(* IEC 61131-3 sources: 2026_Projet_YGO_ExcavatriceDragage/TOOLS/TEST_AUTO_CI/RESULTS/B_AU_SECURITE/reports, 1 file *)

(* ---- FB_Safety_EmergencyManagement_test.st ---- *)
SETUP
VAR
    fb : FB_SAFETY_EMERGENCYMANAGEMENT;
END_VAR
END_SETUP

(* Profil actif : 12 preuves fonctionnelles AF. Les essais de causes et diagnostics sont conserves dans contract_deferred. *)

(* Ordre de rapport stable : contrat IEC, scenarios operationnels, puis TC-P01 par numero croissant. *)

TEST 'TC-P03-001 Dynamique Enable : neutralisation initiale, transition Ready au repos, puis coupure'
    (* Scan 0 : Enable=FALSE -> Neutralisation standard *)
    fb(ENABLE := FALSE, RESET := FALSE, ARMREQUEST := FALSE, POWERCUTOFFREQUEST := FALSE,
       BTNEMERGENCYCUTOFF := FALSE, EMERGENCYCHAINCLOSED := TRUE, POWERCONTACTORENGAGED := FALSE);
    fb(ENABLE := FALSE, RESET := FALSE, ARMREQUEST := FALSE, POWERCUTOFFREQUEST := FALSE,
       BTNEMERGENCYCUTOFF := FALSE, EMERGENCYCHAINCLOSED := TRUE, POWERCONTACTORENGAGED := FALSE);
    ASSERT_FALSE(fb.STATUS.READY, 'Enable=FALSE -> Ready=FALSE (neutralise)');
    ASSERT_FALSE(fb.STATUS.DIAG.ERROR, 'Enable=FALSE -> Pas d erreur');
    ASSERT_FALSE(fb.CMD.MAINTAINA_CMD, 'Enable=FALSE -> MaintainA_Cmd=FALSE (projection fail-safe §10)');
    ASSERT_FALSE(fb.CMD.MAINTAINB_CMD, 'Enable=FALSE -> MaintainB_Cmd=FALSE (projection fail-safe §10)');
    ASSERT_FALSE(fb.CMD.ARMPULSE_CMD, 'Enable=FALSE -> ArmPulse_Cmd=FALSE (projection fail-safe §10)');
    ASSERT_EQ(fb.STATUS.STATE.STEP, 0, 'Enable=FALSE -> sequence neutralisee, Step=0');
    ASSERT_EQ(fb.STATUS.OPERATORMESSAGE, 'AU neutralisee (Enable=FALSE)', 'message neutralisation (gate §2, priorite §11)');

    ADVANCE_TIME(10000000);

    (* Scan 1 : Enable=TRUE -> Prete en service *)
    fb(ENABLE := TRUE, RESET := FALSE, ARMREQUEST := FALSE, POWERCUTOFFREQUEST := FALSE,
       BTNEMERGENCYCUTOFF := FALSE, EMERGENCYCHAINCLOSED := TRUE, POWERCONTACTORENGAGED := FALSE);
    fb(ENABLE := TRUE, RESET := FALSE, ARMREQUEST := FALSE, POWERCUTOFFREQUEST := FALSE,
       BTNEMERGENCYCUTOFF := FALSE, EMERGENCYCHAINCLOSED := TRUE, POWERCONTACTORENGAGED := FALSE);
    ASSERT_TRUE(fb.STATUS.READY, 'Enable=TRUE -> Ready=TRUE (nominal)');
    ASSERT_FALSE(fb.STATUS.DIAG.ERROR, 'Au repos -> Pas d erreur');

    ADVANCE_TIME(10000000);

    (* Scan 2 : Enable=FALSE -> Re-neutralisation *)
    fb(ENABLE := FALSE, RESET := FALSE, ARMREQUEST := FALSE, POWERCUTOFFREQUEST := FALSE,
       BTNEMERGENCYCUTOFF := FALSE, EMERGENCYCHAINCLOSED := TRUE, POWERCONTACTORENGAGED := FALSE);
    fb(ENABLE := FALSE, RESET := FALSE, ARMREQUEST := FALSE, POWERCUTOFFREQUEST := FALSE,
       BTNEMERGENCYCUTOFF := FALSE, EMERGENCYCHAINCLOSED := TRUE, POWERCONTACTORENGAGED := FALSE);
    ASSERT_FALSE(fb.STATUS.READY, 'Coupure -> Ready retombe a FALSE');
END_TEST

TEST 'TC-P01-SCEN-NOM Scenario Nominal : Sequence complete de rearmement sans blocage'
    (* 💤 Étape 0 : Repos initial (machine hors tension, contacteur au repos, Armable=TRUE) *)
    fb(ENABLE := TRUE, RESET := FALSE, ARMREQUEST := FALSE, POWERCUTOFFREQUEST := FALSE,
       BTNEMERGENCYCUTOFF := FALSE, EMERGENCYCHAINCLOSED := TRUE, POWERCONTACTORENGAGED := FALSE);
    fb(ENABLE := TRUE, RESET := FALSE, ARMREQUEST := FALSE, POWERCUTOFFREQUEST := FALSE,
       BTNEMERGENCYCUTOFF := FALSE, EMERGENCYCHAINCLOSED := TRUE, POWERCONTACTORENGAGED := FALSE);
    ADVANCE_TIME(10000000);
    fb(ENABLE := TRUE, RESET := FALSE, ARMREQUEST := FALSE, POWERCUTOFFREQUEST := FALSE,
       BTNEMERGENCYCUTOFF := FALSE, EMERGENCYCHAINCLOSED := TRUE, POWERCONTACTORENGAGED := FALSE);
    fb(ENABLE := TRUE, RESET := FALSE, ARMREQUEST := FALSE, POWERCUTOFFREQUEST := FALSE,
       BTNEMERGENCYCUTOFF := FALSE, EMERGENCYCHAINCLOSED := TRUE, POWERCONTACTORENGAGED := FALSE);
    ASSERT_TRUE(fb.STATUS.STATE.ARMABLE, 'Au repos boucle saine -> Armable=TRUE');
    ASSERT_FALSE(fb.STATUS.DONE, 'Puissance non encore engagee -> Done=FALSE');
    ASSERT_EQ(fb.STATUS.OPERATORMESSAGE, 'AU: repos - pret a rearmer', 'message CASE 0/IDLE au repos sain');

    (* ⏱️ Étape 0bis : Demande de réarmement (Front ArmRequest -> Délai pré-armement 500ms en Step 0) *)
    ADVANCE_TIME(10000000);
    fb(ENABLE := TRUE, RESET := FALSE, ARMREQUEST := TRUE, POWERCUTOFFREQUEST := FALSE,
       BTNEMERGENCYCUTOFF := FALSE, EMERGENCYCHAINCLOSED := TRUE, POWERCONTACTORENGAGED := FALSE);
    fb(ENABLE := TRUE, RESET := FALSE, ARMREQUEST := TRUE, POWERCUTOFFREQUEST := FALSE,
       BTNEMERGENCYCUTOFF := FALSE, EMERGENCYCHAINCLOSED := TRUE, POWERCONTACTORENGAGED := FALSE);
    ASSERT_EQ(fb.STATUS.STATE.STEP, 0, 'Front ArmRequest lance delai pre-armement (reste Step 0)');
    ASSERT_EQ(fb.STATUS.OPERATORMESSAGE, 'AU: appui pris en compte - etablissement chaine', 'message pre-armement actif');

    (* 🚀 Étape 1 : Écoulement 500ms -> Entrée en TestA (Step 1, durée 1s) *)
    ADVANCE_TIME(500000000);
    fb(ENABLE := TRUE, RESET := FALSE, ARMREQUEST := FALSE, POWERCUTOFFREQUEST := FALSE,
       BTNEMERGENCYCUTOFF := FALSE, EMERGENCYCHAINCLOSED := TRUE, POWERCONTACTORENGAGED := FALSE);
    fb(ENABLE := TRUE, RESET := FALSE, ARMREQUEST := FALSE, POWERCUTOFFREQUEST := FALSE,
       BTNEMERGENCYCUTOFF := FALSE, EMERGENCYCHAINCLOSED := TRUE, POWERCONTACTORENGAGED := FALSE);
    ASSERT_EQ(fb.STATUS.STATE.STEP, 1, 'Delai 500ms ecoule -> Entree en TestA');
    ASSERT_EQ(fb.STATUS.OPERATORMESSAGE, 'AU: autotest canal A en cours', 'message CASE 1/TEST_A');
    ASSERT_FALSE(fb.CMD.MAINTAINA_CMD, 'TestA coupe canal A');
    ASSERT_TRUE(fb.CMD.MAINTAINB_CMD, 'TestA maintient canal B');

    (* 🔍 Étape 2 : Écoulement 1s TestA + réaction boucle -> Passage à RestoreA (500ms settle) *)
    ADVANCE_TIME(1000000000);
    fb(ENABLE := TRUE, RESET := FALSE, ARMREQUEST := FALSE, POWERCUTOFFREQUEST := FALSE,
       BTNEMERGENCYCUTOFF := FALSE, EMERGENCYCHAINCLOSED := FALSE, POWERCONTACTORENGAGED := FALSE);
    fb(ENABLE := TRUE, RESET := FALSE, ARMREQUEST := FALSE, POWERCUTOFFREQUEST := FALSE,
       BTNEMERGENCYCUTOFF := FALSE, EMERGENCYCHAINCLOSED := FALSE, POWERCONTACTORENGAGED := FALSE);
    ASSERT_EQ(fb.STATUS.STATE.STEP, 2, 'TestA 1s ecoule + boucle tombee -> RestoreA');
    ASSERT_TRUE(fb.CMD.MAINTAINA_CMD, 'Canal A restaure');
    ASSERT_TRUE(fb.CMD.MAINTAINB_CMD, 'Canal B maintenu');

    (* 🔍 Étape 3 : Écoulement 500ms RestoreA + refermeture boucle -> Passage à TestB (1s) *)
    ADVANCE_TIME(500000000);
    fb(ENABLE := TRUE, RESET := FALSE, ARMREQUEST := FALSE, POWERCUTOFFREQUEST := FALSE,
       BTNEMERGENCYCUTOFF := FALSE, EMERGENCYCHAINCLOSED := TRUE, POWERCONTACTORENGAGED := FALSE);
    fb(ENABLE := TRUE, RESET := FALSE, ARMREQUEST := FALSE, POWERCUTOFFREQUEST := FALSE,
       BTNEMERGENCYCUTOFF := FALSE, EMERGENCYCHAINCLOSED := TRUE, POWERCONTACTORENGAGED := FALSE);
    ASSERT_EQ(fb.STATUS.STATE.STEP, 3, 'RestoreA 500ms ecoule + boucle fermee -> TestB');
    ASSERT_EQ(fb.STATUS.OPERATORMESSAGE, 'AU: autotest canal B en cours', 'message CASE 3/TEST_B');
    ASSERT_FALSE(fb.CMD.MAINTAINB_CMD, 'TestB coupe canal B');
    ASSERT_TRUE(fb.CMD.MAINTAINA_CMD, 'TestB maintient canal A');

    (* 🔍 Étape 4 : Écoulement 1s TestB + réaction boucle -> Passage à RestoreB (1s hold) *)
    ADVANCE_TIME(1000000000);
    fb(ENABLE := TRUE, RESET := FALSE, ARMREQUEST := FALSE, POWERCUTOFFREQUEST := FALSE,
       BTNEMERGENCYCUTOFF := FALSE, EMERGENCYCHAINCLOSED := FALSE, POWERCONTACTORENGAGED := FALSE);
    fb(ENABLE := TRUE, RESET := FALSE, ARMREQUEST := FALSE, POWERCUTOFFREQUEST := FALSE,
       BTNEMERGENCYCUTOFF := FALSE, EMERGENCYCHAINCLOSED := FALSE, POWERCONTACTORENGAGED := FALSE);
    ASSERT_EQ(fb.STATUS.STATE.STEP, 4, 'TestB 1s ecoule + boucle tombee -> RestoreB');
    ASSERT_TRUE(fb.CMD.MAINTAINB_CMD, 'Canal B restaure');
    ASSERT_TRUE(fb.CMD.MAINTAINA_CMD, 'Canal A maintenu');

    (* ⚡ Étape 5 : Écoulement 1s RestoreB (KeepAliveHold) + boucle refermée -> Step 5 Impulsion 1s *)
    ADVANCE_TIME(1000000000);
    fb(ENABLE := TRUE, RESET := FALSE, ARMREQUEST := FALSE, POWERCUTOFFREQUEST := FALSE,
       BTNEMERGENCYCUTOFF := FALSE, EMERGENCYCHAINCLOSED := TRUE, POWERCONTACTORENGAGED := FALSE);
    fb(ENABLE := TRUE, RESET := FALSE, ARMREQUEST := FALSE, POWERCUTOFFREQUEST := FALSE,
       BTNEMERGENCYCUTOFF := FALSE, EMERGENCYCHAINCLOSED := TRUE, POWERCONTACTORENGAGED := FALSE);
    ASSERT_EQ(fb.STATUS.STATE.STEP, 5, 'Auto-test A/B valide -> Step 5 Impulsion contacteur');
    ASSERT_EQ(fb.STATUS.OPERATORMESSAGE, 'AU: impulsion rearmement contacteur', 'message CASE 5/PULSE');
    ASSERT_TRUE(fb.CMD.ARMPULSE_CMD, 'Impulsion 1s active');

    (* ⏱️ Étape 6 : Écoulement 1s impulsion -> Attente confirmation contacteur (Step 6) *)
    ADVANCE_TIME(1000000000);
    fb(ENABLE := TRUE, RESET := FALSE, ARMREQUEST := FALSE, POWERCUTOFFREQUEST := FALSE,
       BTNEMERGENCYCUTOFF := FALSE, EMERGENCYCHAINCLOSED := TRUE, POWERCONTACTORENGAGED := FALSE);
    fb(ENABLE := TRUE, RESET := FALSE, ARMREQUEST := FALSE, POWERCUTOFFREQUEST := FALSE,
       BTNEMERGENCYCUTOFF := FALSE, EMERGENCYCHAINCLOSED := TRUE, POWERCONTACTORENGAGED := FALSE);
    ASSERT_EQ(fb.STATUS.STATE.STEP, 6, 'Impulsion terminee -> Step 6 Confirmation');
    ASSERT_EQ(fb.STATUS.OPERATORMESSAGE, 'AU: attente confirmation contacteur', 'message CASE 6/CONFIRM');
    ASSERT_FALSE(fb.CMD.ARMPULSE_CMD, 'Impulsion retombe');

    (* ✅ Étape 7 : Confirmation contacteur engagé -> Puissance engagée & Latch WasArmed *)
    ADVANCE_TIME(10000000);
    fb(ENABLE := TRUE, RESET := FALSE, ARMREQUEST := FALSE, POWERCUTOFFREQUEST := FALSE,
       BTNEMERGENCYCUTOFF := FALSE, EMERGENCYCHAINCLOSED := TRUE, POWERCONTACTORENGAGED := TRUE);
    fb(ENABLE := TRUE, RESET := FALSE, ARMREQUEST := FALSE, POWERCUTOFFREQUEST := FALSE,
       BTNEMERGENCYCUTOFF := FALSE, EMERGENCYCHAINCLOSED := TRUE, POWERCONTACTORENGAGED := TRUE);
    ASSERT_EQ(fb.STATUS.STATE.STEP, 0, 'Contacteur confirme -> Retour repos IDLE');
    ASSERT_TRUE(fb.STATUS.DONE, 'Puissance engagee -> Done=TRUE');
    ASSERT_TRUE(fb.STATUS.DIAG.WASARMED, 'WasArmed latche a TRUE');
    ASSERT_FALSE(fb.STATUS.DIAG.ERROR, 'Cycle nominal termine sans defaut');
END_TEST

TEST 'TC-P01-SCEN-DYN Scenario Dynamique : Enchainement nominal puis perturbations reelles en service'
    (* 🚀 Phase 1 : Réarmement nominal réussi et mise en service *)
    fb(ENABLE := TRUE, RESET := FALSE, ARMREQUEST := FALSE, POWERCUTOFFREQUEST := FALSE,
       BTNEMERGENCYCUTOFF := FALSE, EMERGENCYCHAINCLOSED := TRUE, POWERCONTACTORENGAGED := FALSE);
    fb(ENABLE := TRUE, RESET := FALSE, ARMREQUEST := FALSE, POWERCUTOFFREQUEST := FALSE,
       BTNEMERGENCYCUTOFF := FALSE, EMERGENCYCHAINCLOSED := TRUE, POWERCONTACTORENGAGED := FALSE);
    ADVANCE_TIME(10000000);
    fb(ENABLE := TRUE, RESET := FALSE, ARMREQUEST := TRUE, POWERCUTOFFREQUEST := FALSE,
       BTNEMERGENCYCUTOFF := FALSE, EMERGENCYCHAINCLOSED := TRUE, POWERCONTACTORENGAGED := FALSE);
    fb(ENABLE := TRUE, RESET := FALSE, ARMREQUEST := TRUE, POWERCUTOFFREQUEST := FALSE,
       BTNEMERGENCYCUTOFF := FALSE, EMERGENCYCHAINCLOSED := TRUE, POWERCONTACTORENGAGED := FALSE);
    ADVANCE_TIME(500000000); // 500ms pre-arm
    fb(ENABLE := TRUE, RESET := FALSE, ARMREQUEST := FALSE, POWERCUTOFFREQUEST := FALSE,
       BTNEMERGENCYCUTOFF := FALSE, EMERGENCYCHAINCLOSED := TRUE, POWERCONTACTORENGAGED := FALSE);
    fb(ENABLE := TRUE, RESET := FALSE, ARMREQUEST := FALSE, POWERCUTOFFREQUEST := FALSE,
       BTNEMERGENCYCUTOFF := FALSE, EMERGENCYCHAINCLOSED := TRUE, POWERCONTACTORENGAGED := FALSE);
    ADVANCE_TIME(1000000000); // 1s TestA
    fb(ENABLE := TRUE, RESET := FALSE, ARMREQUEST := FALSE, POWERCUTOFFREQUEST := FALSE,
       BTNEMERGENCYCUTOFF := FALSE, EMERGENCYCHAINCLOSED := FALSE, POWERCONTACTORENGAGED := FALSE);
    fb(ENABLE := TRUE, RESET := FALSE, ARMREQUEST := FALSE, POWERCUTOFFREQUEST := FALSE,
       BTNEMERGENCYCUTOFF := FALSE, EMERGENCYCHAINCLOSED := FALSE, POWERCONTACTORENGAGED := FALSE);
    ADVANCE_TIME(500000000); // 500ms RestoreA
    fb(ENABLE := TRUE, RESET := FALSE, ARMREQUEST := FALSE, POWERCUTOFFREQUEST := FALSE,
       BTNEMERGENCYCUTOFF := FALSE, EMERGENCYCHAINCLOSED := TRUE, POWERCONTACTORENGAGED := FALSE);
    fb(ENABLE := TRUE, RESET := FALSE, ARMREQUEST := FALSE, POWERCUTOFFREQUEST := FALSE,
       BTNEMERGENCYCUTOFF := FALSE, EMERGENCYCHAINCLOSED := TRUE, POWERCONTACTORENGAGED := FALSE);
    ADVANCE_TIME(1000000000); // 1s TestB
    fb(ENABLE := TRUE, RESET := FALSE, ARMREQUEST := FALSE, POWERCUTOFFREQUEST := FALSE,
       BTNEMERGENCYCUTOFF := FALSE, EMERGENCYCHAINCLOSED := FALSE, POWERCONTACTORENGAGED := FALSE);
    fb(ENABLE := TRUE, RESET := FALSE, ARMREQUEST := FALSE, POWERCUTOFFREQUEST := FALSE,
       BTNEMERGENCYCUTOFF := FALSE, EMERGENCYCHAINCLOSED := FALSE, POWERCONTACTORENGAGED := FALSE);
    ADVANCE_TIME(1000000000); // 1s RestoreB
    fb(ENABLE := TRUE, RESET := FALSE, ARMREQUEST := FALSE, POWERCUTOFFREQUEST := FALSE,
       BTNEMERGENCYCUTOFF := FALSE, EMERGENCYCHAINCLOSED := TRUE, POWERCONTACTORENGAGED := FALSE);
    fb(ENABLE := TRUE, RESET := FALSE, ARMREQUEST := FALSE, POWERCUTOFFREQUEST := FALSE,
       BTNEMERGENCYCUTOFF := FALSE, EMERGENCYCHAINCLOSED := TRUE, POWERCONTACTORENGAGED := FALSE);
    ADVANCE_TIME(1000000000); // 1s Pulse
    fb(ENABLE := TRUE, RESET := FALSE, ARMREQUEST := FALSE, POWERCUTOFFREQUEST := FALSE,
       BTNEMERGENCYCUTOFF := FALSE, EMERGENCYCHAINCLOSED := TRUE, POWERCONTACTORENGAGED := FALSE);
    fb(ENABLE := TRUE, RESET := FALSE, ARMREQUEST := FALSE, POWERCUTOFFREQUEST := FALSE,
       BTNEMERGENCYCUTOFF := FALSE, EMERGENCYCHAINCLOSED := TRUE, POWERCONTACTORENGAGED := FALSE);
    ADVANCE_TIME(10000000);
    fb(ENABLE := TRUE, RESET := FALSE, ARMREQUEST := FALSE, POWERCUTOFFREQUEST := FALSE,
       BTNEMERGENCYCUTOFF := FALSE, EMERGENCYCHAINCLOSED := TRUE, POWERCONTACTORENGAGED := TRUE);
    fb(ENABLE := TRUE, RESET := FALSE, ARMREQUEST := FALSE, POWERCUTOFFREQUEST := FALSE,
       BTNEMERGENCYCUTOFF := FALSE, EMERGENCYCHAINCLOSED := TRUE, POWERCONTACTORENGAGED := TRUE);
    ASSERT_TRUE(fb.STATUS.DONE, 'Machine armee en service');

    (* ⚡ Phase 2 : Coupure sécurité métier intempestive en pleine marche *)
    ADVANCE_TIME(500000000);
    fb(ENABLE := TRUE, RESET := FALSE, ARMREQUEST := FALSE, POWERCUTOFFREQUEST := TRUE,
       BTNEMERGENCYCUTOFF := FALSE, EMERGENCYCHAINCLOSED := TRUE, POWERCONTACTORENGAGED := FALSE);
    fb(ENABLE := TRUE, RESET := FALSE, ARMREQUEST := FALSE, POWERCUTOFFREQUEST := TRUE,
       BTNEMERGENCYCUTOFF := FALSE, EMERGENCYCHAINCLOSED := TRUE, POWERCONTACTORENGAGED := FALSE);
    ASSERT_FALSE(fb.CMD.MAINTAINA_CMD, 'Coupure metier -> Retombee immediate canal A');
    ASSERT_FALSE(fb.CMD.MAINTAINB_CMD, 'Coupure metier -> Retombee immediate canal B');
    ASSERT_FALSE(fb.STATUS.STATE.ARMABLE, 'Coupure metier active -> Armable=FALSE');

    (* 🛡️ Phase 3 : Tentative de réarmement bloquée sous défaut *)
    ADVANCE_TIME(10000000);
    fb(ENABLE := TRUE, RESET := FALSE, ARMREQUEST := TRUE, POWERCUTOFFREQUEST := TRUE,
       BTNEMERGENCYCUTOFF := FALSE, EMERGENCYCHAINCLOSED := TRUE, POWERCONTACTORENGAGED := FALSE);
    fb(ENABLE := TRUE, RESET := FALSE, ARMREQUEST := TRUE, POWERCUTOFFREQUEST := TRUE,
       BTNEMERGENCYCUTOFF := FALSE, EMERGENCYCHAINCLOSED := TRUE, POWERCONTACTORENGAGED := FALSE);
    ASSERT_EQ(fb.STATUS.STATE.STEP, 0, 'Rearmement refuse : reste a Step 0');

    (* 🔄 Phase 4 : Disparition de la dérive métier + écoulement garde 5s + Acquittement Reset *)
    ADVANCE_TIME(5000000000); // écoulement 5s garde anti-chatter
    fb(ENABLE := TRUE, RESET := TRUE, ARMREQUEST := FALSE, POWERCUTOFFREQUEST := FALSE,
       BTNEMERGENCYCUTOFF := FALSE, EMERGENCYCHAINCLOSED := TRUE, POWERCONTACTORENGAGED := FALSE);
    fb(ENABLE := TRUE, RESET := TRUE, ARMREQUEST := FALSE, POWERCUTOFFREQUEST := FALSE,
       BTNEMERGENCYCUTOFF := FALSE, EMERGENCYCHAINCLOSED := TRUE, POWERCONTACTORENGAGED := FALSE);
    ASSERT_TRUE(fb.STATUS.STATE.ARMABLE, 'Defaut acquitte et disparu -> Armable redevient TRUE');

    (* ⚠️ Phase 5 : Nouvel armement avec échec de collage contacteur (timeout 2s) *)
    ADVANCE_TIME(10000000);
    fb(ENABLE := TRUE, RESET := FALSE, ARMREQUEST := TRUE, POWERCUTOFFREQUEST := FALSE,
       BTNEMERGENCYCUTOFF := FALSE, EMERGENCYCHAINCLOSED := TRUE, POWERCONTACTORENGAGED := FALSE);
    fb(ENABLE := TRUE, RESET := FALSE, ARMREQUEST := TRUE, POWERCUTOFFREQUEST := FALSE,
       BTNEMERGENCYCUTOFF := FALSE, EMERGENCYCHAINCLOSED := TRUE, POWERCONTACTORENGAGED := FALSE);
    ADVANCE_TIME(500000000); // 500ms pre-arm
    fb(ENABLE := TRUE, RESET := FALSE, ARMREQUEST := FALSE, POWERCUTOFFREQUEST := FALSE,
       BTNEMERGENCYCUTOFF := FALSE, EMERGENCYCHAINCLOSED := TRUE, POWERCONTACTORENGAGED := FALSE);
    fb(ENABLE := TRUE, RESET := FALSE, ARMREQUEST := FALSE, POWERCUTOFFREQUEST := FALSE,
       BTNEMERGENCYCUTOFF := FALSE, EMERGENCYCHAINCLOSED := TRUE, POWERCONTACTORENGAGED := FALSE);
    ADVANCE_TIME(1000000000); // 1s TestA
    fb(ENABLE := TRUE, RESET := FALSE, ARMREQUEST := FALSE, POWERCUTOFFREQUEST := FALSE,
       BTNEMERGENCYCUTOFF := FALSE, EMERGENCYCHAINCLOSED := FALSE, POWERCONTACTORENGAGED := FALSE);
    fb(ENABLE := TRUE, RESET := FALSE, ARMREQUEST := FALSE, POWERCUTOFFREQUEST := FALSE,
       BTNEMERGENCYCUTOFF := FALSE, EMERGENCYCHAINCLOSED := FALSE, POWERCONTACTORENGAGED := FALSE);
    ADVANCE_TIME(500000000); // 500ms RestoreA
    fb(ENABLE := TRUE, RESET := FALSE, ARMREQUEST := FALSE, POWERCUTOFFREQUEST := FALSE,
       BTNEMERGENCYCUTOFF := FALSE, EMERGENCYCHAINCLOSED := TRUE, POWERCONTACTORENGAGED := FALSE);
    fb(ENABLE := TRUE, RESET := FALSE, ARMREQUEST := FALSE, POWERCUTOFFREQUEST := FALSE,
       BTNEMERGENCYCUTOFF := FALSE, EMERGENCYCHAINCLOSED := TRUE, POWERCONTACTORENGAGED := FALSE);
    ADVANCE_TIME(1000000000); // 1s TestB
    fb(ENABLE := TRUE, RESET := FALSE, ARMREQUEST := FALSE, POWERCUTOFFREQUEST := FALSE,
       BTNEMERGENCYCUTOFF := FALSE, EMERGENCYCHAINCLOSED := FALSE, POWERCONTACTORENGAGED := FALSE);
    fb(ENABLE := TRUE, RESET := FALSE, ARMREQUEST := FALSE, POWERCUTOFFREQUEST := FALSE,
       BTNEMERGENCYCUTOFF := FALSE, EMERGENCYCHAINCLOSED := FALSE, POWERCONTACTORENGAGED := FALSE);
    ADVANCE_TIME(1000000000); // 1s RestoreB
    fb(ENABLE := TRUE, RESET := FALSE, ARMREQUEST := FALSE, POWERCUTOFFREQUEST := FALSE,
       BTNEMERGENCYCUTOFF := FALSE, EMERGENCYCHAINCLOSED := TRUE, POWERCONTACTORENGAGED := FALSE);
    fb(ENABLE := TRUE, RESET := FALSE, ARMREQUEST := FALSE, POWERCUTOFFREQUEST := FALSE,
       BTNEMERGENCYCUTOFF := FALSE, EMERGENCYCHAINCLOSED := TRUE, POWERCONTACTORENGAGED := FALSE);
    ADVANCE_TIME(1000000000); // 1s Pulse
    fb(ENABLE := TRUE, RESET := FALSE, ARMREQUEST := FALSE, POWERCUTOFFREQUEST := FALSE,
       BTNEMERGENCYCUTOFF := FALSE, EMERGENCYCHAINCLOSED := TRUE, POWERCONTACTORENGAGED := FALSE);
    fb(ENABLE := TRUE, RESET := FALSE, ARMREQUEST := FALSE, POWERCUTOFFREQUEST := FALSE,
       BTNEMERGENCYCUTOFF := FALSE, EMERGENCYCHAINCLOSED := TRUE, POWERCONTACTORENGAGED := FALSE);

    (* Timeout 2s à l'étape 6 sans retour PowerContactorEngaged *)
    ADVANCE_TIME(2000000000);
    fb(ENABLE := TRUE, RESET := FALSE, ARMREQUEST := FALSE, POWERCUTOFFREQUEST := FALSE,
       BTNEMERGENCYCUTOFF := FALSE, EMERGENCYCHAINCLOSED := TRUE, POWERCONTACTORENGAGED := FALSE);
    fb(ENABLE := TRUE, RESET := FALSE, ARMREQUEST := FALSE, POWERCUTOFFREQUEST := FALSE,
       BTNEMERGENCYCUTOFF := FALSE, EMERGENCYCHAINCLOSED := TRUE, POWERCONTACTORENGAGED := FALSE);
    ASSERT_TRUE(fb.STATUS.DIAG.ERROR, 'Echec collage contacteur -> Alarme levee');
    ASSERT_TRUE(fb.STATUS.DIAG.LOCKOUTACTIVE, 'Verrouillage Lockout 5s active');
    ASSERT_FALSE(fb.STATUS.STATE.ARMABLE, 'Pendant lockout -> Armable=FALSE');

    (* 🔓 Phase 6 : Expiration du lockout 5s + Reset -> Prêt pour nouvel essai *)
    ADVANCE_TIME(5000000000);
    fb(ENABLE := TRUE, RESET := TRUE, ARMREQUEST := FALSE, POWERCUTOFFREQUEST := FALSE,
       BTNEMERGENCYCUTOFF := FALSE, EMERGENCYCHAINCLOSED := TRUE, POWERCONTACTORENGAGED := FALSE);
    fb(ENABLE := TRUE, RESET := TRUE, ARMREQUEST := FALSE, POWERCUTOFFREQUEST := FALSE,
       BTNEMERGENCYCUTOFF := FALSE, EMERGENCYCHAINCLOSED := TRUE, POWERCONTACTORENGAGED := FALSE);
    ASSERT_FALSE(fb.STATUS.DIAG.LOCKOUTACTIVE, 'Lockout 5s expire');
    ASSERT_TRUE(fb.STATUS.STATE.ARMABLE, 'Machine prete a etre reessayee');
END_TEST

TEST 'TC-P01-001 Coupure AU physique (essai site, non automatise)'
    (* 🟢 SITE — essai terrain, non automatisable en logiciel.
       Enfoncement du coup de poing AU physique sur site -> ouverture materielle
       immediate de la boucle 24V de securite -> retombee instantanee du contacteur
       de puissance ligne (API reste sous tension).
       Maintien PLC : si WasArmed=FALSE, MaintainA/B retombent ; si WasArmed=TRUE,
       les sorties PowerKeepAlive sont preservees (latch WasArmed). *)
    fb(ENABLE := TRUE, RESET := FALSE, ARMREQUEST := FALSE, POWERCUTOFFREQUEST := FALSE,
       BTNEMERGENCYCUTOFF := FALSE, EMERGENCYCHAINCLOSED := FALSE, POWERCONTACTORENGAGED := FALSE);
    fb(ENABLE := TRUE, RESET := FALSE, ARMREQUEST := FALSE, POWERCUTOFFREQUEST := FALSE,
       BTNEMERGENCYCUTOFF := FALSE, EMERGENCYCHAINCLOSED := FALSE, POWERCONTACTORENGAGED := FALSE);
    ASSERT_TRUE(fb.STATUS.STATE.ARMABLE, 'machine hors tension au repos -> Armable=TRUE (rearmement possible)');
    ASSERT_FALSE(fb.CMD.MAINTAINA_CMD, 'avant tout armement (WasArmed=FALSE), maintien canal A retombe');
    ASSERT_FALSE(fb.CMD.MAINTAINB_CMD, 'avant tout armement (WasArmed=FALSE), maintien canal B retombe');
END_TEST

TEST 'TC-P01-002 (partie AUTO) chaque canal est commande independamment, l autre reste maintenu'
    (* demarrage + regime etabli, sain *)
    fb(ENABLE := TRUE, RESET := FALSE, ARMREQUEST := FALSE, POWERCUTOFFREQUEST := FALSE,
       BTNEMERGENCYCUTOFF := FALSE, EMERGENCYCHAINCLOSED := TRUE, POWERCONTACTORENGAGED := FALSE);
    fb(ENABLE := TRUE, RESET := FALSE, ARMREQUEST := FALSE, POWERCUTOFFREQUEST := FALSE,
       BTNEMERGENCYCUTOFF := FALSE, EMERGENCYCHAINCLOSED := TRUE, POWERCONTACTORENGAGED := FALSE);
    ADVANCE_TIME(10000000);
    fb(ENABLE := TRUE, RESET := FALSE, ARMREQUEST := FALSE, POWERCUTOFFREQUEST := FALSE,
       BTNEMERGENCYCUTOFF := FALSE, EMERGENCYCHAINCLOSED := TRUE, POWERCONTACTORENGAGED := FALSE);
    fb(ENABLE := TRUE, RESET := FALSE, ARMREQUEST := FALSE, POWERCUTOFFREQUEST := FALSE,
       BTNEMERGENCYCUTOFF := FALSE, EMERGENCYCHAINCLOSED := TRUE, POWERCONTACTORENGAGED := FALSE);
    ASSERT_TRUE(fb.CMD.MAINTAINA_CMD, 'hors defaut, canal A maintenu');
    ASSERT_TRUE(fb.CMD.MAINTAINB_CMD, 'hors defaut, canal B maintenu');

    (* front ArmRequest -> délai 500ms pre-arm puis TestA (step 1) : SEUL le canal A doit se couper *)
    ADVANCE_TIME(10000000);
    fb(ENABLE := TRUE, RESET := FALSE, ARMREQUEST := TRUE, POWERCUTOFFREQUEST := FALSE,
       BTNEMERGENCYCUTOFF := FALSE, EMERGENCYCHAINCLOSED := TRUE, POWERCONTACTORENGAGED := FALSE);
    fb(ENABLE := TRUE, RESET := FALSE, ARMREQUEST := TRUE, POWERCUTOFFREQUEST := FALSE,
       BTNEMERGENCYCUTOFF := FALSE, EMERGENCYCHAINCLOSED := TRUE, POWERCONTACTORENGAGED := FALSE);
    ADVANCE_TIME(500000000); // 500ms pre-arm
    fb(ENABLE := TRUE, RESET := FALSE, ARMREQUEST := FALSE, POWERCUTOFFREQUEST := FALSE,
       BTNEMERGENCYCUTOFF := FALSE, EMERGENCYCHAINCLOSED := TRUE, POWERCONTACTORENGAGED := FALSE);
    fb(ENABLE := TRUE, RESET := FALSE, ARMREQUEST := FALSE, POWERCUTOFFREQUEST := FALSE,
       BTNEMERGENCYCUTOFF := FALSE, EMERGENCYCHAINCLOSED := TRUE, POWERCONTACTORENGAGED := FALSE);
    ASSERT_EQ(fb.STATUS.STATE.STEP, 1, 'front doit lancer TestA');
    ASSERT_FALSE(fb.CMD.MAINTAINA_CMD, 'TestA : canal A seul doit se couper');
    ASSERT_TRUE(fb.CMD.MAINTAINB_CMD, 'TestA : canal B ne doit PAS etre affecte');

    (* 1s plus tard : la boucle reagit reellement a la coupure de A (preuve physique reelle) *)
    ADVANCE_TIME(1000000000); // 1s TestA
    fb(ENABLE := TRUE, RESET := FALSE, ARMREQUEST := FALSE, POWERCUTOFFREQUEST := FALSE,
       BTNEMERGENCYCUTOFF := FALSE, EMERGENCYCHAINCLOSED := FALSE, POWERCONTACTORENGAGED := FALSE);
    fb(ENABLE := TRUE, RESET := FALSE, ARMREQUEST := FALSE, POWERCUTOFFREQUEST := FALSE,
       BTNEMERGENCYCUTOFF := FALSE, EMERGENCYCHAINCLOSED := FALSE, POWERCONTACTORENGAGED := FALSE);
    ASSERT_EQ(fb.STATUS.STATE.STEP, 2, 'TestA reussi (boucle a reagi) -> RestoreA');
    ASSERT_FALSE(fb.STATUS.DIAG.ERROR, 'pas de defaut si le canal reagit correctement au test');
    ASSERT_TRUE(fb.CMD.MAINTAINA_CMD, 'canal A restaure immediatement apres son test');

    (* 500ms plus tard : boucle refermee (A restaure) -> passage a TestB (step 3) *)
    ADVANCE_TIME(500000000); // 500ms RestoreA
    fb(ENABLE := TRUE, RESET := FALSE, ARMREQUEST := FALSE, POWERCUTOFFREQUEST := FALSE,
       BTNEMERGENCYCUTOFF := FALSE, EMERGENCYCHAINCLOSED := TRUE, POWERCONTACTORENGAGED := FALSE);
    fb(ENABLE := TRUE, RESET := FALSE, ARMREQUEST := FALSE, POWERCUTOFFREQUEST := FALSE,
       BTNEMERGENCYCUTOFF := FALSE, EMERGENCYCHAINCLOSED := TRUE, POWERCONTACTORENGAGED := FALSE);
    ASSERT_EQ(fb.STATUS.STATE.STEP, 3, 'RestoreA reussi -> TestB');
    ASSERT_FALSE(fb.CMD.MAINTAINB_CMD, 'TestB : canal B seul doit se couper');
    ASSERT_TRUE(fb.CMD.MAINTAINA_CMD, 'TestB : canal A ne doit PAS etre affecte');

    (* 1s plus tard : boucle reagit a la coupure de B *)
    ADVANCE_TIME(1000000000); // 1s TestB
    fb(ENABLE := TRUE, RESET := FALSE, ARMREQUEST := FALSE, POWERCUTOFFREQUEST := FALSE,
       BTNEMERGENCYCUTOFF := FALSE, EMERGENCYCHAINCLOSED := FALSE, POWERCONTACTORENGAGED := FALSE);
    fb(ENABLE := TRUE, RESET := FALSE, ARMREQUEST := FALSE, POWERCUTOFFREQUEST := FALSE,
       BTNEMERGENCYCUTOFF := FALSE, EMERGENCYCHAINCLOSED := FALSE, POWERCONTACTORENGAGED := FALSE);
    ASSERT_EQ(fb.STATUS.STATE.STEP, 4, 'TestB reussi -> RestoreB');
    ASSERT_FALSE(fb.STATUS.DIAG.ERROR, 'pas de defaut si le canal B reagit correctement au test');
    ASSERT_TRUE(fb.CMD.MAINTAINB_CMD, 'canal B restaure immediatement apres son test');
END_TEST

TEST 'TC-P01-003 front ArmRequest + boucle OK sur les 2 canaux -> pulse 1s puis confirmation'
    (* demarrage + regime etabli, sain *)
    fb(ENABLE := TRUE, RESET := FALSE, ARMREQUEST := FALSE, POWERCUTOFFREQUEST := FALSE,
       BTNEMERGENCYCUTOFF := FALSE, EMERGENCYCHAINCLOSED := TRUE, POWERCONTACTORENGAGED := FALSE);
    fb(ENABLE := TRUE, RESET := FALSE, ARMREQUEST := FALSE, POWERCUTOFFREQUEST := FALSE,
       BTNEMERGENCYCUTOFF := FALSE, EMERGENCYCHAINCLOSED := TRUE, POWERCONTACTORENGAGED := FALSE);
    ADVANCE_TIME(10000000);
    fb(ENABLE := TRUE, RESET := FALSE, ARMREQUEST := FALSE, POWERCUTOFFREQUEST := FALSE,
       BTNEMERGENCYCUTOFF := FALSE, EMERGENCYCHAINCLOSED := TRUE, POWERCONTACTORENGAGED := FALSE);
    fb(ENABLE := TRUE, RESET := FALSE, ARMREQUEST := FALSE, POWERCUTOFFREQUEST := FALSE,
       BTNEMERGENCYCUTOFF := FALSE, EMERGENCYCHAINCLOSED := TRUE, POWERCONTACTORENGAGED := FALSE);

    (* front ArmRequest -> delai 500ms -> TestA *)
    ADVANCE_TIME(10000000);
    fb(ENABLE := TRUE, RESET := FALSE, ARMREQUEST := TRUE, POWERCUTOFFREQUEST := FALSE,
       BTNEMERGENCYCUTOFF := FALSE, EMERGENCYCHAINCLOSED := TRUE, POWERCONTACTORENGAGED := FALSE);
    fb(ENABLE := TRUE, RESET := FALSE, ARMREQUEST := TRUE, POWERCUTOFFREQUEST := FALSE,
       BTNEMERGENCYCUTOFF := FALSE, EMERGENCYCHAINCLOSED := TRUE, POWERCONTACTORENGAGED := FALSE);
    ADVANCE_TIME(500000000); // 500ms pre-arm
    fb(ENABLE := TRUE, RESET := FALSE, ARMREQUEST := FALSE, POWERCUTOFFREQUEST := FALSE,
       BTNEMERGENCYCUTOFF := FALSE, EMERGENCYCHAINCLOSED := TRUE, POWERCONTACTORENGAGED := FALSE);
    fb(ENABLE := TRUE, RESET := FALSE, ARMREQUEST := FALSE, POWERCUTOFFREQUEST := FALSE,
       BTNEMERGENCYCUTOFF := FALSE, EMERGENCYCHAINCLOSED := TRUE, POWERCONTACTORENGAGED := FALSE);

    (* TestA reussi (boucle reagit) -> RestoreA *)
    ADVANCE_TIME(1000000000); // 1s TestA
    fb(ENABLE := TRUE, RESET := FALSE, ARMREQUEST := FALSE, POWERCUTOFFREQUEST := FALSE,
       BTNEMERGENCYCUTOFF := FALSE, EMERGENCYCHAINCLOSED := FALSE, POWERCONTACTORENGAGED := FALSE);
    fb(ENABLE := TRUE, RESET := FALSE, ARMREQUEST := FALSE, POWERCUTOFFREQUEST := FALSE,
       BTNEMERGENCYCUTOFF := FALSE, EMERGENCYCHAINCLOSED := FALSE, POWERCONTACTORENGAGED := FALSE);

    (* RestoreA reussi -> TestB *)
    ADVANCE_TIME(500000000); // 500ms RestoreA
    fb(ENABLE := TRUE, RESET := FALSE, ARMREQUEST := FALSE, POWERCUTOFFREQUEST := FALSE,
       BTNEMERGENCYCUTOFF := FALSE, EMERGENCYCHAINCLOSED := TRUE, POWERCONTACTORENGAGED := FALSE);
    fb(ENABLE := TRUE, RESET := FALSE, ARMREQUEST := FALSE, POWERCUTOFFREQUEST := FALSE,
       BTNEMERGENCYCUTOFF := FALSE, EMERGENCYCHAINCLOSED := TRUE, POWERCONTACTORENGAGED := FALSE);

    (* TestB reussi (boucle reagit) -> RestoreB *)
    ADVANCE_TIME(1000000000); // 1s TestB
    fb(ENABLE := TRUE, RESET := FALSE, ARMREQUEST := FALSE, POWERCUTOFFREQUEST := FALSE,
       BTNEMERGENCYCUTOFF := FALSE, EMERGENCYCHAINCLOSED := FALSE, POWERCONTACTORENGAGED := FALSE);
    fb(ENABLE := TRUE, RESET := FALSE, ARMREQUEST := FALSE, POWERCUTOFFREQUEST := FALSE,
       BTNEMERGENCYCUTOFF := FALSE, EMERGENCYCHAINCLOSED := FALSE, POWERCONTACTORENGAGED := FALSE);

    (* RestoreB reussi -> Pulse (step 5), impulsion 1s *)
    ADVANCE_TIME(1000000000); // 1s RestoreB
    fb(ENABLE := TRUE, RESET := FALSE, ARMREQUEST := FALSE, POWERCUTOFFREQUEST := FALSE,
       BTNEMERGENCYCUTOFF := FALSE, EMERGENCYCHAINCLOSED := TRUE, POWERCONTACTORENGAGED := FALSE);
    fb(ENABLE := TRUE, RESET := FALSE, ARMREQUEST := FALSE, POWERCUTOFFREQUEST := FALSE,
       BTNEMERGENCYCUTOFF := FALSE, EMERGENCYCHAINCLOSED := TRUE, POWERCONTACTORENGAGED := FALSE);
    ASSERT_EQ(fb.STATUS.STATE.STEP, 5, 'les 2 canaux valides -> impulsion de reamement');
    ASSERT_TRUE(fb.CMD.ARMPULSE_CMD, 'pulse de reamement doit etre actif (TC-P01-003)');

    (* 1s plus tard : pulse termine -> Confirm (step 6) *)
    ADVANCE_TIME(1000000000);
    fb(ENABLE := TRUE, RESET := FALSE, ARMREQUEST := FALSE, POWERCUTOFFREQUEST := FALSE,
       BTNEMERGENCYCUTOFF := FALSE, EMERGENCYCHAINCLOSED := TRUE, POWERCONTACTORENGAGED := FALSE);
    fb(ENABLE := TRUE, RESET := FALSE, ARMREQUEST := FALSE, POWERCUTOFFREQUEST := FALSE,
       BTNEMERGENCYCUTOFF := FALSE, EMERGENCYCHAINCLOSED := TRUE, POWERCONTACTORENGAGED := FALSE);
    ASSERT_EQ(fb.STATUS.STATE.STEP, 6, 'pulse de 1s termine -> attente confirmation contacteur');
    ASSERT_FALSE(fb.CMD.ARMPULSE_CMD, 'pulse retombe apres 1s');
    ASSERT_TRUE(fb.STATUS.STATE.ARMINGBUSY, 'sequence toujours en cours (attente confirmation)');

    (* contacteur confirme engage -> succes, retour IDLE *)
    ADVANCE_TIME(10000000);
    fb(ENABLE := TRUE, RESET := FALSE, ARMREQUEST := FALSE, POWERCUTOFFREQUEST := FALSE,
       BTNEMERGENCYCUTOFF := FALSE, EMERGENCYCHAINCLOSED := TRUE, POWERCONTACTORENGAGED := TRUE);
    fb(ENABLE := TRUE, RESET := FALSE, ARMREQUEST := FALSE, POWERCUTOFFREQUEST := FALSE,
       BTNEMERGENCYCUTOFF := FALSE, EMERGENCYCHAINCLOSED := TRUE, POWERCONTACTORENGAGED := TRUE);
    ASSERT_EQ(fb.STATUS.STATE.STEP, 0, 'confirmation contacteur -> retour IDLE');
    ASSERT_TRUE(fb.STATUS.DONE, 'contacteur engage confirme -> Done');
    ASSERT_FALSE(fb.STATUS.STATE.ARMINGBUSY, 'sequence terminee');
    ASSERT_FALSE(fb.STATUS.DIAG.LOCKOUTACTIVE, 'succes -> pas de lockout');
    ASSERT_FALSE(fb.STATUS.DIAG.ERROR, 'reamement reussi -> pas de defaut');
END_TEST

TEST 'TC-P01-004/009 Reset acquitte l affichage mais re-alarme si la cause persiste'
    (* reproduit l etat "canal colle" de TC-P01-006 -- setup independant, propre a ce test *)
    fb(ENABLE := TRUE, RESET := FALSE, ARMREQUEST := FALSE, POWERCUTOFFREQUEST := FALSE,
       BTNEMERGENCYCUTOFF := FALSE, EMERGENCYCHAINCLOSED := TRUE, POWERCONTACTORENGAGED := FALSE);
    fb(ENABLE := TRUE, RESET := FALSE, ARMREQUEST := FALSE, POWERCUTOFFREQUEST := FALSE,
       BTNEMERGENCYCUTOFF := FALSE, EMERGENCYCHAINCLOSED := TRUE, POWERCONTACTORENGAGED := FALSE);
    ADVANCE_TIME(10000000);
    fb(ENABLE := TRUE, RESET := FALSE, ARMREQUEST := FALSE, POWERCUTOFFREQUEST := FALSE,
       BTNEMERGENCYCUTOFF := FALSE, EMERGENCYCHAINCLOSED := TRUE, POWERCONTACTORENGAGED := FALSE);
    fb(ENABLE := TRUE, RESET := FALSE, ARMREQUEST := FALSE, POWERCUTOFFREQUEST := FALSE,
       BTNEMERGENCYCUTOFF := FALSE, EMERGENCYCHAINCLOSED := TRUE, POWERCONTACTORENGAGED := FALSE);
    ADVANCE_TIME(10000000);
    fb(ENABLE := TRUE, RESET := FALSE, ARMREQUEST := TRUE, POWERCUTOFFREQUEST := FALSE,
       BTNEMERGENCYCUTOFF := FALSE, EMERGENCYCHAINCLOSED := TRUE, POWERCONTACTORENGAGED := FALSE);
    fb(ENABLE := TRUE, RESET := FALSE, ARMREQUEST := TRUE, POWERCUTOFFREQUEST := FALSE,
       BTNEMERGENCYCUTOFF := FALSE, EMERGENCYCHAINCLOSED := TRUE, POWERCONTACTORENGAGED := FALSE);
    ADVANCE_TIME(500000000); // 500ms pre-arm
    fb(ENABLE := TRUE, RESET := FALSE, ARMREQUEST := FALSE, POWERCUTOFFREQUEST := FALSE,
       BTNEMERGENCYCUTOFF := FALSE, EMERGENCYCHAINCLOSED := TRUE, POWERCONTACTORENGAGED := FALSE);
    fb(ENABLE := TRUE, RESET := FALSE, ARMREQUEST := FALSE, POWERCUTOFFREQUEST := FALSE,
       BTNEMERGENCYCUTOFF := FALSE, EMERGENCYCHAINCLOSED := TRUE, POWERCONTACTORENGAGED := FALSE);
    ADVANCE_TIME(1000000000); // 1s TestA avec boucle qui reste fermee (collage)
    fb(ENABLE := TRUE, RESET := FALSE, ARMREQUEST := FALSE, POWERCUTOFFREQUEST := FALSE,
       BTNEMERGENCYCUTOFF := FALSE, EMERGENCYCHAINCLOSED := TRUE, POWERCONTACTORENGAGED := FALSE);
    fb(ENABLE := TRUE, RESET := FALSE, ARMREQUEST := FALSE, POWERCUTOFFREQUEST := FALSE,
       BTNEMERGENCYCUTOFF := FALSE, EMERGENCYCHAINCLOSED := TRUE, POWERCONTACTORENGAGED := FALSE);
    ASSERT_TRUE(fb.STATUS.DIAG.ERROR, 'precondition : canal colle doit avoir leve une erreur');

    (* Reset : doit acquitter l affichage sans redemarrage auto (TC-P01-004) -- +1 cycle *)
    ADVANCE_TIME(10000000);
    fb(ENABLE := TRUE, RESET := TRUE, ARMREQUEST := FALSE, POWERCUTOFFREQUEST := FALSE,
       BTNEMERGENCYCUTOFF := FALSE, EMERGENCYCHAINCLOSED := TRUE, POWERCONTACTORENGAGED := FALSE);
    fb(ENABLE := TRUE, RESET := TRUE, ARMREQUEST := FALSE, POWERCUTOFFREQUEST := FALSE,
       BTNEMERGENCYCUTOFF := FALSE, EMERGENCYCHAINCLOSED := TRUE, POWERCONTACTORENGAGED := FALSE);
    ASSERT_FALSE(fb.STATUS.DIAG.ERROR, 'Reset doit effacer l affichage du defaut');
    ASSERT_EQ(fb.STATUS.STATE.STEP, 0, 'Reset seul ne relance jamais de sequence (pas de redemarrage auto)');
    ASSERT_TRUE(fb.CMD.MAINTAINA_CMD, 'Reset acquitte la cause redondance figee -> maintien autorise hors defaut');

    (* Ecoulement de la garde 5s anti-chatter avant de retenter un front *)
    ADVANCE_TIME(5000000000);
    fb(ENABLE := TRUE, RESET := FALSE, ARMREQUEST := FALSE, POWERCUTOFFREQUEST := FALSE,
       BTNEMERGENCYCUTOFF := FALSE, EMERGENCYCHAINCLOSED := TRUE, POWERCONTACTORENGAGED := FALSE);
    fb(ENABLE := TRUE, RESET := FALSE, ARMREQUEST := FALSE, POWERCUTOFFREQUEST := FALSE,
       BTNEMERGENCYCUTOFF := FALSE, EMERGENCYCHAINCLOSED := TRUE, POWERCONTACTORENGAGED := FALSE);

    (* nouvel essai : cause toujours presente (canal toujours colle) -> doit re-alarmer (TC-P01-009) *)
    ADVANCE_TIME(10000000);
    fb(ENABLE := TRUE, RESET := FALSE, ARMREQUEST := TRUE, POWERCUTOFFREQUEST := FALSE,
       BTNEMERGENCYCUTOFF := FALSE, EMERGENCYCHAINCLOSED := TRUE, POWERCONTACTORENGAGED := FALSE);
    fb(ENABLE := TRUE, RESET := FALSE, ARMREQUEST := TRUE, POWERCUTOFFREQUEST := FALSE,
       BTNEMERGENCYCUTOFF := FALSE, EMERGENCYCHAINCLOSED := TRUE, POWERCONTACTORENGAGED := FALSE);
    ADVANCE_TIME(500000000); // 500ms pre-arm -> lance TestA
    fb(ENABLE := TRUE, RESET := FALSE, ARMREQUEST := FALSE, POWERCUTOFFREQUEST := FALSE,
       BTNEMERGENCYCUTOFF := FALSE, EMERGENCYCHAINCLOSED := TRUE, POWERCONTACTORENGAGED := FALSE);
    fb(ENABLE := TRUE, RESET := FALSE, ARMREQUEST := FALSE, POWERCUTOFFREQUEST := FALSE,
       BTNEMERGENCYCUTOFF := FALSE, EMERGENCYCHAINCLOSED := TRUE, POWERCONTACTORENGAGED := FALSE);
    ASSERT_EQ(fb.STATUS.STATE.STEP, 1, 'un nouveau front ArmRequest doit relancer TestA');

    ADVANCE_TIME(1000000000); // 1s TestA canal colle
    fb(ENABLE := TRUE, RESET := FALSE, ARMREQUEST := FALSE, POWERCUTOFFREQUEST := FALSE,
       BTNEMERGENCYCUTOFF := FALSE, EMERGENCYCHAINCLOSED := TRUE, POWERCONTACTORENGAGED := FALSE);
    fb(ENABLE := TRUE, RESET := FALSE, ARMREQUEST := FALSE, POWERCUTOFFREQUEST := FALSE,
       BTNEMERGENCYCUTOFF := FALSE, EMERGENCYCHAINCLOSED := TRUE, POWERCONTACTORENGAGED := FALSE);
    ASSERT_TRUE(fb.STATUS.DIAG.ERROR, 'cause persistante doit re-alarmer au nouvel essai, meme apres Reset');
END_TEST

TEST 'TC-P01-005 Sequence 2 temps : ArmRequest sans Reset bloque ; Reset puis ArmRequest arme'
    (* Setup : montee en sequence jusqu au pulse (steps 1-5), puis timeout confirmation 2s
       -> EmergencyArmingFailed + lockout 5s *)
    fb(ENABLE := TRUE, RESET := FALSE, ARMREQUEST := FALSE, POWERCUTOFFREQUEST := FALSE,
       BTNEMERGENCYCUTOFF := FALSE, EMERGENCYCHAINCLOSED := TRUE, POWERCONTACTORENGAGED := FALSE);
    fb(ENABLE := TRUE, RESET := FALSE, ARMREQUEST := FALSE, POWERCUTOFFREQUEST := FALSE,
       BTNEMERGENCYCUTOFF := FALSE, EMERGENCYCHAINCLOSED := TRUE, POWERCONTACTORENGAGED := FALSE);
    ADVANCE_TIME(10000000);
    fb(ENABLE := TRUE, RESET := FALSE, ARMREQUEST := FALSE, POWERCUTOFFREQUEST := FALSE,
       BTNEMERGENCYCUTOFF := FALSE, EMERGENCYCHAINCLOSED := TRUE, POWERCONTACTORENGAGED := FALSE);
    fb(ENABLE := TRUE, RESET := FALSE, ARMREQUEST := FALSE, POWERCUTOFFREQUEST := FALSE,
       BTNEMERGENCYCUTOFF := FALSE, EMERGENCYCHAINCLOSED := TRUE, POWERCONTACTORENGAGED := FALSE);
    ADVANCE_TIME(10000000);
    fb(ENABLE := TRUE, RESET := FALSE, ARMREQUEST := TRUE, POWERCUTOFFREQUEST := FALSE,
       BTNEMERGENCYCUTOFF := FALSE, EMERGENCYCHAINCLOSED := TRUE, POWERCONTACTORENGAGED := FALSE);
    fb(ENABLE := TRUE, RESET := FALSE, ARMREQUEST := TRUE, POWERCUTOFFREQUEST := FALSE,
       BTNEMERGENCYCUTOFF := FALSE, EMERGENCYCHAINCLOSED := TRUE, POWERCONTACTORENGAGED := FALSE);
    ADVANCE_TIME(500000000); // 500ms pre-arm
    fb(ENABLE := TRUE, RESET := FALSE, ARMREQUEST := FALSE, POWERCUTOFFREQUEST := FALSE,
       BTNEMERGENCYCUTOFF := FALSE, EMERGENCYCHAINCLOSED := TRUE, POWERCONTACTORENGAGED := FALSE);
    fb(ENABLE := TRUE, RESET := FALSE, ARMREQUEST := FALSE, POWERCUTOFFREQUEST := FALSE,
       BTNEMERGENCYCUTOFF := FALSE, EMERGENCYCHAINCLOSED := TRUE, POWERCONTACTORENGAGED := FALSE);
    ADVANCE_TIME(1000000000); // 1s TestA
    fb(ENABLE := TRUE, RESET := FALSE, ARMREQUEST := FALSE, POWERCUTOFFREQUEST := FALSE,
       BTNEMERGENCYCUTOFF := FALSE, EMERGENCYCHAINCLOSED := FALSE, POWERCONTACTORENGAGED := FALSE);
    fb(ENABLE := TRUE, RESET := FALSE, ARMREQUEST := FALSE, POWERCUTOFFREQUEST := FALSE,
       BTNEMERGENCYCUTOFF := FALSE, EMERGENCYCHAINCLOSED := FALSE, POWERCONTACTORENGAGED := FALSE);
    ADVANCE_TIME(500000000); // 500ms RestoreA
    fb(ENABLE := TRUE, RESET := FALSE, ARMREQUEST := FALSE, POWERCUTOFFREQUEST := FALSE,
       BTNEMERGENCYCUTOFF := FALSE, EMERGENCYCHAINCLOSED := TRUE, POWERCONTACTORENGAGED := FALSE);
    fb(ENABLE := TRUE, RESET := FALSE, ARMREQUEST := FALSE, POWERCUTOFFREQUEST := FALSE,
       BTNEMERGENCYCUTOFF := FALSE, EMERGENCYCHAINCLOSED := TRUE, POWERCONTACTORENGAGED := FALSE);
    ADVANCE_TIME(1000000000); // 1s TestB
    fb(ENABLE := TRUE, RESET := FALSE, ARMREQUEST := FALSE, POWERCUTOFFREQUEST := FALSE,
       BTNEMERGENCYCUTOFF := FALSE, EMERGENCYCHAINCLOSED := FALSE, POWERCONTACTORENGAGED := FALSE);
    fb(ENABLE := TRUE, RESET := FALSE, ARMREQUEST := FALSE, POWERCUTOFFREQUEST := FALSE,
       BTNEMERGENCYCUTOFF := FALSE, EMERGENCYCHAINCLOSED := FALSE, POWERCONTACTORENGAGED := FALSE);
    ADVANCE_TIME(1000000000); // 1s RestoreB
    fb(ENABLE := TRUE, RESET := FALSE, ARMREQUEST := FALSE, POWERCUTOFFREQUEST := FALSE,
       BTNEMERGENCYCUTOFF := FALSE, EMERGENCYCHAINCLOSED := TRUE, POWERCONTACTORENGAGED := FALSE);
    fb(ENABLE := TRUE, RESET := FALSE, ARMREQUEST := FALSE, POWERCUTOFFREQUEST := FALSE,
       BTNEMERGENCYCUTOFF := FALSE, EMERGENCYCHAINCLOSED := TRUE, POWERCONTACTORENGAGED := FALSE);
    ADVANCE_TIME(1000000000); // 1s Pulse
    fb(ENABLE := TRUE, RESET := FALSE, ARMREQUEST := FALSE, POWERCUTOFFREQUEST := FALSE,
       BTNEMERGENCYCUTOFF := FALSE, EMERGENCYCHAINCLOSED := TRUE, POWERCONTACTORENGAGED := FALSE);
    fb(ENABLE := TRUE, RESET := FALSE, ARMREQUEST := FALSE, POWERCUTOFFREQUEST := FALSE,
       BTNEMERGENCYCUTOFF := FALSE, EMERGENCYCHAINCLOSED := TRUE, POWERCONTACTORENGAGED := FALSE);
    (* timeout 2s confirmation -> EmergencyArmingFailed + lockout *)
    ADVANCE_TIME(2000000000);
    fb(ENABLE := TRUE, RESET := FALSE, ARMREQUEST := FALSE, POWERCUTOFFREQUEST := FALSE,
       BTNEMERGENCYCUTOFF := FALSE, EMERGENCYCHAINCLOSED := TRUE, POWERCONTACTORENGAGED := FALSE);
    fb(ENABLE := TRUE, RESET := FALSE, ARMREQUEST := FALSE, POWERCUTOFFREQUEST := FALSE,
       BTNEMERGENCYCUTOFF := FALSE, EMERGENCYCHAINCLOSED := TRUE, POWERCONTACTORENGAGED := FALSE);
    ASSERT_TRUE(fb.STATUS.DIAG.LOCKOUTACTIVE, 'precondition : lockout 5s actif apres echec');
    ASSERT_FALSE(fb.STATUS.STATE.ARMABLE, 'precondition : Armable=FALSE sous lockout');

    (* Temps 1 : ArmRequest SANS Reset -> bloque (lockout actif), reste Step 0 *)
    ADVANCE_TIME(10000000);
    fb(ENABLE := TRUE, RESET := FALSE, ARMREQUEST := TRUE, POWERCUTOFFREQUEST := FALSE,
       BTNEMERGENCYCUTOFF := FALSE, EMERGENCYCHAINCLOSED := TRUE, POWERCONTACTORENGAGED := FALSE);
    fb(ENABLE := TRUE, RESET := FALSE, ARMREQUEST := TRUE, POWERCUTOFFREQUEST := FALSE,
       BTNEMERGENCYCUTOFF := FALSE, EMERGENCYCHAINCLOSED := TRUE, POWERCONTACTORENGAGED := FALSE);
    ASSERT_EQ(fb.STATUS.STATE.STEP, 0, 'Temps 1 : ArmRequest sans Reset bloque -> reste Step 0');

    (* Temps 2a : Reset acquitte et purge le defaut + lockout *)
    ADVANCE_TIME(10000000);
    fb(ENABLE := TRUE, RESET := TRUE, ARMREQUEST := FALSE, POWERCUTOFFREQUEST := FALSE,
       BTNEMERGENCYCUTOFF := FALSE, EMERGENCYCHAINCLOSED := TRUE, POWERCONTACTORENGAGED := FALSE);
    fb(ENABLE := TRUE, RESET := TRUE, ARMREQUEST := FALSE, POWERCUTOFFREQUEST := FALSE,
       BTNEMERGENCYCUTOFF := FALSE, EMERGENCYCHAINCLOSED := TRUE, POWERCONTACTORENGAGED := FALSE);
    ASSERT_FALSE(fb.STATUS.DIAG.LOCKOUTACTIVE, 'Reset purge le lockout');
    ASSERT_FALSE(fb.STATUS.DIAG.ERROR, 'Reset acquitte l affichage du defaut');

    (* Ecoulement garde anti-chatter *)
    ADVANCE_TIME(5000000000);
    fb(ENABLE := TRUE, RESET := FALSE, ARMREQUEST := FALSE, POWERCUTOFFREQUEST := FALSE,
       BTNEMERGENCYCUTOFF := FALSE, EMERGENCYCHAINCLOSED := TRUE, POWERCONTACTORENGAGED := FALSE);
    fb(ENABLE := TRUE, RESET := FALSE, ARMREQUEST := FALSE, POWERCUTOFFREQUEST := FALSE,
       BTNEMERGENCYCUTOFF := FALSE, EMERGENCYCHAINCLOSED := TRUE, POWERCONTACTORENGAGED := FALSE);

    (* Temps 2b : ArmRequest distinct et conscient -> délai 500ms -> arme (Step 1) *)
    ADVANCE_TIME(10000000);
    fb(ENABLE := TRUE, RESET := FALSE, ARMREQUEST := TRUE, POWERCUTOFFREQUEST := FALSE,
       BTNEMERGENCYCUTOFF := FALSE, EMERGENCYCHAINCLOSED := TRUE, POWERCONTACTORENGAGED := FALSE);
    fb(ENABLE := TRUE, RESET := FALSE, ARMREQUEST := TRUE, POWERCUTOFFREQUEST := FALSE,
       BTNEMERGENCYCUTOFF := FALSE, EMERGENCYCHAINCLOSED := TRUE, POWERCONTACTORENGAGED := FALSE);
    ADVANCE_TIME(500000000); // 500ms pre-arm
    fb(ENABLE := TRUE, RESET := FALSE, ARMREQUEST := FALSE, POWERCUTOFFREQUEST := FALSE,
       BTNEMERGENCYCUTOFF := FALSE, EMERGENCYCHAINCLOSED := TRUE, POWERCONTACTORENGAGED := FALSE);
    fb(ENABLE := TRUE, RESET := FALSE, ARMREQUEST := FALSE, POWERCUTOFFREQUEST := FALSE,
       BTNEMERGENCYCUTOFF := FALSE, EMERGENCYCHAINCLOSED := TRUE, POWERCONTACTORENGAGED := FALSE);
    ASSERT_EQ(fb.STATUS.STATE.STEP, 1, 'Temps 2 : Reset puis ArmRequest -> sequence armee (Step 1)');
END_TEST

TEST 'TC-P01-006 canal colle bloque le reamement (echec auto-test)'
    (* scans 1-2 : demarrage + regime etabli, sain *)
    fb(ENABLE := TRUE, RESET := FALSE, ARMREQUEST := FALSE, POWERCUTOFFREQUEST := FALSE,
       BTNEMERGENCYCUTOFF := FALSE, EMERGENCYCHAINCLOSED := TRUE, POWERCONTACTORENGAGED := FALSE);
    fb(ENABLE := TRUE, RESET := FALSE, ARMREQUEST := FALSE, POWERCUTOFFREQUEST := FALSE,
       BTNEMERGENCYCUTOFF := FALSE, EMERGENCYCHAINCLOSED := TRUE, POWERCONTACTORENGAGED := FALSE);
    ADVANCE_TIME(10000000);
    fb(ENABLE := TRUE, RESET := FALSE, ARMREQUEST := FALSE, POWERCUTOFFREQUEST := FALSE,
       BTNEMERGENCYCUTOFF := FALSE, EMERGENCYCHAINCLOSED := TRUE, POWERCONTACTORENGAGED := FALSE);
    fb(ENABLE := TRUE, RESET := FALSE, ARMREQUEST := FALSE, POWERCUTOFFREQUEST := FALSE,
       BTNEMERGENCYCUTOFF := FALSE, EMERGENCYCHAINCLOSED := TRUE, POWERCONTACTORENGAGED := FALSE);

    (* front ArmRequest -> delai 500ms -> ArmingSeqStep passe a 1 (TestA) *)
    ADVANCE_TIME(10000000);
    fb(ENABLE := TRUE, RESET := FALSE, ARMREQUEST := TRUE, POWERCUTOFFREQUEST := FALSE,
       BTNEMERGENCYCUTOFF := FALSE, EMERGENCYCHAINCLOSED := TRUE, POWERCONTACTORENGAGED := FALSE);
    fb(ENABLE := TRUE, RESET := FALSE, ARMREQUEST := TRUE, POWERCUTOFFREQUEST := FALSE,
       BTNEMERGENCYCUTOFF := FALSE, EMERGENCYCHAINCLOSED := TRUE, POWERCONTACTORENGAGED := FALSE);
    ADVANCE_TIME(500000000); // 500ms pre-arm
    fb(ENABLE := TRUE, RESET := FALSE, ARMREQUEST := FALSE, POWERCUTOFFREQUEST := FALSE,
       BTNEMERGENCYCUTOFF := FALSE, EMERGENCYCHAINCLOSED := TRUE, POWERCONTACTORENGAGED := FALSE);
    fb(ENABLE := TRUE, RESET := FALSE, ARMREQUEST := FALSE, POWERCUTOFFREQUEST := FALSE,
       BTNEMERGENCYCUTOFF := FALSE, EMERGENCYCHAINCLOSED := TRUE, POWERCONTACTORENGAGED := FALSE);
    ASSERT_EQ(fb.STATUS.STATE.STEP, 1, 'front ArmRequest doit lancer TestA (step 1)');

    (* 1s plus tard : le canal A est cense etre coupe, mais la boucle reste fermee -> collage *)
    ADVANCE_TIME(1000000000); // 1s TestA
    fb(ENABLE := TRUE, RESET := FALSE, ARMREQUEST := FALSE, POWERCUTOFFREQUEST := FALSE,
       BTNEMERGENCYCUTOFF := FALSE, EMERGENCYCHAINCLOSED := TRUE, POWERCONTACTORENGAGED := FALSE);
    fb(ENABLE := TRUE, RESET := FALSE, ARMREQUEST := FALSE, POWERCUTOFFREQUEST := FALSE,
       BTNEMERGENCYCUTOFF := FALSE, EMERGENCYCHAINCLOSED := TRUE, POWERCONTACTORENGAGED := FALSE);
    ASSERT_TRUE(fb.STATUS.DIAG.ERROR, 'canal colle doit lever une erreur (RedundancyTestFailed)');
    ASSERT_EQ(fb.STATUS.OPERATORMESSAGE, 'AU: defaut redondance contacteurs - verifier puis Reset', 'message defaut redondance');
    ASSERT_EQ(fb.STATUS.STATE.STEP, 0, 'echec auto-test doit ramener la sequence a IDLE');
    ASSERT_FALSE(fb.CMD.MAINTAINA_CMD, 'un canal colle bloque aussi le maintien normal (interlock sur Cause brute)');
    ASSERT_EQ(fb.STATUS.DIAG.LASTABORTSTEP, 1, 'abandon a l etape 1 (TestA)');
    ASSERT_EQ(fb.STATUS.DIAG.LASTABORTCAUSE, 16#0020, 'cause = 16#0020 (CST_ABORT_REDUNDANCY_A = 32)');
    ASSERT_TRUE(fb.STATUS.DIAG.REDUNDANCYTESTFAILED, 'defaut redondance leve (Diag.RedundancyTestFailed)');
    ASSERT_FALSE(fb.CMD.MAINTAINB_CMD, 'canal colle bloque aussi le maintien B (interlock Cause brute sur les 2 canaux)');
END_TEST

TEST 'TC-P01-007 timeout confirmation contacteur -> lockout 5s'
    (* meme montee en sequence que TC-P01-003 : les 2 canaux valides, jusqu au pulse *)
    fb(ENABLE := TRUE, RESET := FALSE, ARMREQUEST := FALSE, POWERCUTOFFREQUEST := FALSE,
       BTNEMERGENCYCUTOFF := FALSE, EMERGENCYCHAINCLOSED := TRUE, POWERCONTACTORENGAGED := FALSE);
    fb(ENABLE := TRUE, RESET := FALSE, ARMREQUEST := FALSE, POWERCUTOFFREQUEST := FALSE,
       BTNEMERGENCYCUTOFF := FALSE, EMERGENCYCHAINCLOSED := TRUE, POWERCONTACTORENGAGED := FALSE);
    ADVANCE_TIME(10000000);
    fb(ENABLE := TRUE, RESET := FALSE, ARMREQUEST := FALSE, POWERCUTOFFREQUEST := FALSE,
       BTNEMERGENCYCUTOFF := FALSE, EMERGENCYCHAINCLOSED := TRUE, POWERCONTACTORENGAGED := FALSE);
    fb(ENABLE := TRUE, RESET := FALSE, ARMREQUEST := FALSE, POWERCUTOFFREQUEST := FALSE,
       BTNEMERGENCYCUTOFF := FALSE, EMERGENCYCHAINCLOSED := TRUE, POWERCONTACTORENGAGED := FALSE);
    ADVANCE_TIME(10000000);
    fb(ENABLE := TRUE, RESET := FALSE, ARMREQUEST := TRUE, POWERCUTOFFREQUEST := FALSE,
       BTNEMERGENCYCUTOFF := FALSE, EMERGENCYCHAINCLOSED := TRUE, POWERCONTACTORENGAGED := FALSE);
    fb(ENABLE := TRUE, RESET := FALSE, ARMREQUEST := TRUE, POWERCUTOFFREQUEST := FALSE,
       BTNEMERGENCYCUTOFF := FALSE, EMERGENCYCHAINCLOSED := TRUE, POWERCONTACTORENGAGED := FALSE);
    ADVANCE_TIME(500000000); // 500ms pre-arm
    fb(ENABLE := TRUE, RESET := FALSE, ARMREQUEST := FALSE, POWERCUTOFFREQUEST := FALSE,
       BTNEMERGENCYCUTOFF := FALSE, EMERGENCYCHAINCLOSED := TRUE, POWERCONTACTORENGAGED := FALSE);
    fb(ENABLE := TRUE, RESET := FALSE, ARMREQUEST := FALSE, POWERCUTOFFREQUEST := FALSE,
       BTNEMERGENCYCUTOFF := FALSE, EMERGENCYCHAINCLOSED := TRUE, POWERCONTACTORENGAGED := FALSE);
    ADVANCE_TIME(1000000000); // 1s TestA
    fb(ENABLE := TRUE, RESET := FALSE, ARMREQUEST := FALSE, POWERCUTOFFREQUEST := FALSE,
       BTNEMERGENCYCUTOFF := FALSE, EMERGENCYCHAINCLOSED := FALSE, POWERCONTACTORENGAGED := FALSE);
    fb(ENABLE := TRUE, RESET := FALSE, ARMREQUEST := FALSE, POWERCUTOFFREQUEST := FALSE,
       BTNEMERGENCYCUTOFF := FALSE, EMERGENCYCHAINCLOSED := FALSE, POWERCONTACTORENGAGED := FALSE);
    ADVANCE_TIME(500000000); // 500ms RestoreA
    fb(ENABLE := TRUE, RESET := FALSE, ARMREQUEST := FALSE, POWERCUTOFFREQUEST := FALSE,
       BTNEMERGENCYCUTOFF := FALSE, EMERGENCYCHAINCLOSED := TRUE, POWERCONTACTORENGAGED := FALSE);
    fb(ENABLE := TRUE, RESET := FALSE, ARMREQUEST := FALSE, POWERCUTOFFREQUEST := FALSE,
       BTNEMERGENCYCUTOFF := FALSE, EMERGENCYCHAINCLOSED := TRUE, POWERCONTACTORENGAGED := FALSE);
    ADVANCE_TIME(1000000000); // 1s TestB
    fb(ENABLE := TRUE, RESET := FALSE, ARMREQUEST := FALSE, POWERCUTOFFREQUEST := FALSE,
       BTNEMERGENCYCUTOFF := FALSE, EMERGENCYCHAINCLOSED := FALSE, POWERCONTACTORENGAGED := FALSE);
    fb(ENABLE := TRUE, RESET := FALSE, ARMREQUEST := FALSE, POWERCUTOFFREQUEST := FALSE,
       BTNEMERGENCYCUTOFF := FALSE, EMERGENCYCHAINCLOSED := FALSE, POWERCONTACTORENGAGED := FALSE);
    ADVANCE_TIME(1000000000); // 1s RestoreB
    fb(ENABLE := TRUE, RESET := FALSE, ARMREQUEST := FALSE, POWERCUTOFFREQUEST := FALSE,
       BTNEMERGENCYCUTOFF := FALSE, EMERGENCYCHAINCLOSED := TRUE, POWERCONTACTORENGAGED := FALSE);
    fb(ENABLE := TRUE, RESET := FALSE, ARMREQUEST := FALSE, POWERCUTOFFREQUEST := FALSE,
       BTNEMERGENCYCUTOFF := FALSE, EMERGENCYCHAINCLOSED := TRUE, POWERCONTACTORENGAGED := FALSE);
    ASSERT_EQ(fb.STATUS.STATE.STEP, 5, 'les 2 canaux valides -> pulse');

    (* 1s plus tard : pulse termine -> Confirm (step 6), contacteur PAS engage *)
    ADVANCE_TIME(1000000000);
    fb(ENABLE := TRUE, RESET := FALSE, ARMREQUEST := FALSE, POWERCUTOFFREQUEST := FALSE,
       BTNEMERGENCYCUTOFF := FALSE, EMERGENCYCHAINCLOSED := TRUE, POWERCONTACTORENGAGED := FALSE);
    fb(ENABLE := TRUE, RESET := FALSE, ARMREQUEST := FALSE, POWERCUTOFFREQUEST := FALSE,
       BTNEMERGENCYCUTOFF := FALSE, EMERGENCYCHAINCLOSED := TRUE, POWERCONTACTORENGAGED := FALSE);
    ASSERT_EQ(fb.STATUS.STATE.STEP, 6, 'attente confirmation contacteur');

    (* 2s plus tard (timeout confirmation) : contacteur toujours pas confirme -> echec + lockout *)
    ADVANCE_TIME(2000000000);
    fb(ENABLE := TRUE, RESET := FALSE, ARMREQUEST := FALSE, POWERCUTOFFREQUEST := FALSE,
       BTNEMERGENCYCUTOFF := FALSE, EMERGENCYCHAINCLOSED := TRUE, POWERCONTACTORENGAGED := FALSE);
    fb(ENABLE := TRUE, RESET := FALSE, ARMREQUEST := FALSE, POWERCUTOFFREQUEST := FALSE,
       BTNEMERGENCYCUTOFF := FALSE, EMERGENCYCHAINCLOSED := TRUE, POWERCONTACTORENGAGED := FALSE);
    ASSERT_EQ(fb.STATUS.STATE.STEP, 0, 'timeout confirmation doit ramener la sequence a IDLE');
    ASSERT_EQ(fb.STATUS.DIAG.LASTABORTSTEP, 6, 'abandon a l etape 6 (Confirm)');
    ASSERT_EQ(fb.STATUS.DIAG.LASTABORTCAUSE, 16#0080, 'cause = 16#0080 (CST_ABORT_TIMEOUT_CONTACTOR = 128)');
    ASSERT_EQ(fb.STATUS.OPERATORMESSAGE, 'AU echec: contacteur non confirme', 'message echec rearmement contacteur');
    ASSERT_TRUE(fb.STATUS.DIAG.LOCKOUTACTIVE, 'timeout doit declencher le lockout (TC-P01-007)');
    ASSERT_TRUE(fb.STATUS.DIAG.ARMFAILED, 'timeout doit lever le defaut EmergencyArmingFailed');
    ASSERT_TRUE(fb.STATUS.DIAG.ERROR, 'defaut doit etre visible sur Error');

    (* pendant le lockout : un nouveau front ArmRequest doit etre bloque *)
    ADVANCE_TIME(10000000);
    fb(ENABLE := TRUE, RESET := FALSE, ARMREQUEST := TRUE, POWERCUTOFFREQUEST := FALSE,
       BTNEMERGENCYCUTOFF := FALSE, EMERGENCYCHAINCLOSED := TRUE, POWERCONTACTORENGAGED := FALSE);
    fb(ENABLE := TRUE, RESET := FALSE, ARMREQUEST := TRUE, POWERCUTOFFREQUEST := FALSE,
       BTNEMERGENCYCUTOFF := FALSE, EMERGENCYCHAINCLOSED := TRUE, POWERCONTACTORENGAGED := FALSE);
    ASSERT_EQ(fb.STATUS.STATE.STEP, 0, 'lockout actif doit bloquer toute nouvelle tentative de reamement');

    (* 5s apres le debut du lockout : le verrouillage doit se lever automatiquement *)
    ADVANCE_TIME(5000000000);
    fb(ENABLE := TRUE, RESET := FALSE, ARMREQUEST := FALSE, POWERCUTOFFREQUEST := FALSE,
       BTNEMERGENCYCUTOFF := FALSE, EMERGENCYCHAINCLOSED := TRUE, POWERCONTACTORENGAGED := FALSE);
    fb(ENABLE := TRUE, RESET := FALSE, ARMREQUEST := FALSE, POWERCUTOFFREQUEST := FALSE,
       BTNEMERGENCYCUTOFF := FALSE, EMERGENCYCHAINCLOSED := TRUE, POWERCONTACTORENGAGED := FALSE);
    ASSERT_FALSE(fb.STATUS.DIAG.LOCKOUTACTIVE, 'lockout 5s ecoule -> leve automatiquement');

    (* Reset pour acquitter le defaut *)
    ADVANCE_TIME(10000000);
    fb(ENABLE := TRUE, RESET := TRUE, ARMREQUEST := FALSE, POWERCUTOFFREQUEST := FALSE,
       BTNEMERGENCYCUTOFF := FALSE, EMERGENCYCHAINCLOSED := TRUE, POWERCONTACTORENGAGED := FALSE);
    fb(ENABLE := TRUE, RESET := TRUE, ARMREQUEST := FALSE, POWERCUTOFFREQUEST := FALSE,
       BTNEMERGENCYCUTOFF := FALSE, EMERGENCYCHAINCLOSED := TRUE, POWERCONTACTORENGAGED := FALSE);

    (* nouveau front -> delai 500ms -> relance TestA *)
    ADVANCE_TIME(10000000);
    fb(ENABLE := TRUE, RESET := FALSE, ARMREQUEST := TRUE, POWERCUTOFFREQUEST := FALSE,
       BTNEMERGENCYCUTOFF := FALSE, EMERGENCYCHAINCLOSED := TRUE, POWERCONTACTORENGAGED := FALSE);
    fb(ENABLE := TRUE, RESET := FALSE, ARMREQUEST := TRUE, POWERCUTOFFREQUEST := FALSE,
       BTNEMERGENCYCUTOFF := FALSE, EMERGENCYCHAINCLOSED := TRUE, POWERCONTACTORENGAGED := FALSE);
    ADVANCE_TIME(500000000); // 500ms pre-arm
    fb(ENABLE := TRUE, RESET := FALSE, ARMREQUEST := FALSE, POWERCUTOFFREQUEST := FALSE,
       BTNEMERGENCYCUTOFF := FALSE, EMERGENCYCHAINCLOSED := TRUE, POWERCONTACTORENGAGED := FALSE);
    fb(ENABLE := TRUE, RESET := FALSE, ARMREQUEST := FALSE, POWERCUTOFFREQUEST := FALSE,
       BTNEMERGENCYCUTOFF := FALSE, EMERGENCYCHAINCLOSED := TRUE, POWERCONTACTORENGAGED := FALSE);
    ASSERT_EQ(fb.STATUS.STATE.STEP, 1, 'apres le lockout et Reset, un nouveau front doit relancer TestA');
END_TEST

TEST 'TC-P01-008 PowerCutOffRequest coupe A et B sans armer'
    (* scan 1 : autotest demarrage (1 cycle, boucle saine, contacteur repos) *)
    fb(ENABLE := TRUE, RESET := FALSE, ARMREQUEST := FALSE, POWERCUTOFFREQUEST := FALSE,
       BTNEMERGENCYCUTOFF := FALSE, EMERGENCYCHAINCLOSED := TRUE, POWERCONTACTORENGAGED := FALSE);
    fb(ENABLE := TRUE, RESET := FALSE, ARMREQUEST := FALSE, POWERCUTOFFREQUEST := FALSE,
       BTNEMERGENCYCUTOFF := FALSE, EMERGENCYCHAINCLOSED := TRUE, POWERCONTACTORENGAGED := FALSE);

    (* scan 2 : regime etabli, maintien sain attendu -- +1 cycle automate (10ms) *)
    ADVANCE_TIME(10000000);
    fb(ENABLE := TRUE, RESET := FALSE, ARMREQUEST := FALSE, POWERCUTOFFREQUEST := FALSE,
       BTNEMERGENCYCUTOFF := FALSE, EMERGENCYCHAINCLOSED := TRUE, POWERCONTACTORENGAGED := FALSE);
    fb(ENABLE := TRUE, RESET := FALSE, ARMREQUEST := FALSE, POWERCUTOFFREQUEST := FALSE,
       BTNEMERGENCYCUTOFF := FALSE, EMERGENCYCHAINCLOSED := TRUE, POWERCONTACTORENGAGED := FALSE);
    ASSERT_TRUE(fb.CMD.MAINTAINA_CMD, 'hors defaut, canal A doit etre maintenu');
    ASSERT_TRUE(fb.CMD.MAINTAINB_CMD, 'hors defaut, canal B doit etre maintenu');
    ASSERT_EQ(fb.STATUS.STATE.STEP, 0, 'pas de sequence en cours');

    (* scan 3 : coupure demandee par un metier (Winch/Translation) -- +1 cycle automate *)
    ADVANCE_TIME(10000000);
    fb(ENABLE := TRUE, RESET := FALSE, ARMREQUEST := FALSE, POWERCUTOFFREQUEST := TRUE,
       BTNEMERGENCYCUTOFF := FALSE, EMERGENCYCHAINCLOSED := TRUE, POWERCONTACTORENGAGED := FALSE);
    fb(ENABLE := TRUE, RESET := FALSE, ARMREQUEST := FALSE, POWERCUTOFFREQUEST := TRUE,
       BTNEMERGENCYCUTOFF := FALSE, EMERGENCYCHAINCLOSED := TRUE, POWERCONTACTORENGAGED := FALSE);
    ASSERT_FALSE(fb.CMD.MAINTAINA_CMD, 'PowerCutOffRequest doit couper le canal A');
    ASSERT_FALSE(fb.CMD.MAINTAINB_CMD, 'PowerCutOffRequest doit couper le canal B');
    ASSERT_EQ(fb.STATUS.STATE.STEP, 0, 'PowerCutOffRequest ne doit jamais declencher une sequence armement');
END_TEST

TEST 'TC-P01-010 BtnEmergencyCutOff pendant le pulse de reamement (step 5) doit couper le pulse comme le maintien'
    (* Meme montee en sequence que TC-P01-003 jusqu au pulse (step 5) *)
    fb(ENABLE := TRUE, RESET := FALSE, ARMREQUEST := FALSE, POWERCUTOFFREQUEST := FALSE,
       BTNEMERGENCYCUTOFF := FALSE, EMERGENCYCHAINCLOSED := TRUE, POWERCONTACTORENGAGED := FALSE);
    fb(ENABLE := TRUE, RESET := FALSE, ARMREQUEST := FALSE, POWERCUTOFFREQUEST := FALSE,
       BTNEMERGENCYCUTOFF := FALSE, EMERGENCYCHAINCLOSED := TRUE, POWERCONTACTORENGAGED := FALSE);
    ADVANCE_TIME(10000000);
    fb(ENABLE := TRUE, RESET := FALSE, ARMREQUEST := FALSE, POWERCUTOFFREQUEST := FALSE,
       BTNEMERGENCYCUTOFF := FALSE, EMERGENCYCHAINCLOSED := TRUE, POWERCONTACTORENGAGED := FALSE);
    fb(ENABLE := TRUE, RESET := FALSE, ARMREQUEST := FALSE, POWERCUTOFFREQUEST := FALSE,
       BTNEMERGENCYCUTOFF := FALSE, EMERGENCYCHAINCLOSED := TRUE, POWERCONTACTORENGAGED := FALSE);
    ADVANCE_TIME(10000000);
    fb(ENABLE := TRUE, RESET := FALSE, ARMREQUEST := TRUE, POWERCUTOFFREQUEST := FALSE,
       BTNEMERGENCYCUTOFF := FALSE, EMERGENCYCHAINCLOSED := TRUE, POWERCONTACTORENGAGED := FALSE);
    fb(ENABLE := TRUE, RESET := FALSE, ARMREQUEST := TRUE, POWERCUTOFFREQUEST := FALSE,
       BTNEMERGENCYCUTOFF := FALSE, EMERGENCYCHAINCLOSED := TRUE, POWERCONTACTORENGAGED := FALSE);
    ADVANCE_TIME(500000000); // 500ms pre-arm
    fb(ENABLE := TRUE, RESET := FALSE, ARMREQUEST := FALSE, POWERCUTOFFREQUEST := FALSE,
       BTNEMERGENCYCUTOFF := FALSE, EMERGENCYCHAINCLOSED := TRUE, POWERCONTACTORENGAGED := FALSE);
    fb(ENABLE := TRUE, RESET := FALSE, ARMREQUEST := FALSE, POWERCUTOFFREQUEST := FALSE,
       BTNEMERGENCYCUTOFF := FALSE, EMERGENCYCHAINCLOSED := TRUE, POWERCONTACTORENGAGED := FALSE);
    ADVANCE_TIME(1000000000); // 1s TestA
    fb(ENABLE := TRUE, RESET := FALSE, ARMREQUEST := FALSE, POWERCUTOFFREQUEST := FALSE,
       BTNEMERGENCYCUTOFF := FALSE, EMERGENCYCHAINCLOSED := FALSE, POWERCONTACTORENGAGED := FALSE);
    fb(ENABLE := TRUE, RESET := FALSE, ARMREQUEST := FALSE, POWERCUTOFFREQUEST := FALSE,
       BTNEMERGENCYCUTOFF := FALSE, EMERGENCYCHAINCLOSED := FALSE, POWERCONTACTORENGAGED := FALSE);
    ADVANCE_TIME(500000000); // 500ms RestoreA
    fb(ENABLE := TRUE, RESET := FALSE, ARMREQUEST := FALSE, POWERCUTOFFREQUEST := FALSE,
       BTNEMERGENCYCUTOFF := FALSE, EMERGENCYCHAINCLOSED := TRUE, POWERCONTACTORENGAGED := FALSE);
    fb(ENABLE := TRUE, RESET := FALSE, ARMREQUEST := FALSE, POWERCUTOFFREQUEST := FALSE,
       BTNEMERGENCYCUTOFF := FALSE, EMERGENCYCHAINCLOSED := TRUE, POWERCONTACTORENGAGED := FALSE);
    ADVANCE_TIME(1000000000); // 1s TestB
    fb(ENABLE := TRUE, RESET := FALSE, ARMREQUEST := FALSE, POWERCUTOFFREQUEST := FALSE,
       BTNEMERGENCYCUTOFF := FALSE, EMERGENCYCHAINCLOSED := FALSE, POWERCONTACTORENGAGED := FALSE);
    fb(ENABLE := TRUE, RESET := FALSE, ARMREQUEST := FALSE, POWERCUTOFFREQUEST := FALSE,
       BTNEMERGENCYCUTOFF := FALSE, EMERGENCYCHAINCLOSED := FALSE, POWERCONTACTORENGAGED := FALSE);
    ADVANCE_TIME(1000000000); // 1s RestoreB
    fb(ENABLE := TRUE, RESET := FALSE, ARMREQUEST := FALSE, POWERCUTOFFREQUEST := FALSE,
       BTNEMERGENCYCUTOFF := FALSE, EMERGENCYCHAINCLOSED := TRUE, POWERCONTACTORENGAGED := FALSE);
    fb(ENABLE := TRUE, RESET := FALSE, ARMREQUEST := FALSE, POWERCUTOFFREQUEST := FALSE,
       BTNEMERGENCYCUTOFF := FALSE, EMERGENCYCHAINCLOSED := TRUE, POWERCONTACTORENGAGED := FALSE);
    ASSERT_EQ(fb.STATUS.STATE.STEP, 5, 'les 2 canaux valides -> pulse (step 5)');
    ASSERT_TRUE(fb.CMD.ARMPULSE_CMD, 'precondition : pulse actif');

    (* Operateur appuie sur la coupure d urgence IHM PENDANT l impulsion mecanique de reamement *)
    ADVANCE_TIME(10000000);
    fb(ENABLE := TRUE, RESET := FALSE, ARMREQUEST := FALSE, POWERCUTOFFREQUEST := FALSE,
       BTNEMERGENCYCUTOFF := TRUE, EMERGENCYCHAINCLOSED := TRUE, POWERCONTACTORENGAGED := FALSE);
    fb(ENABLE := TRUE, RESET := FALSE, ARMREQUEST := FALSE, POWERCUTOFFREQUEST := FALSE,
       BTNEMERGENCYCUTOFF := TRUE, EMERGENCYCHAINCLOSED := TRUE, POWERCONTACTORENGAGED := FALSE);
    ASSERT_FALSE(fb.CMD.MAINTAINA_CMD, 'BtnEmergencyCutOff coupe bien le maintien canal A');
    ASSERT_FALSE(fb.CMD.MAINTAINB_CMD, 'BtnEmergencyCutOff coupe bien le maintien canal B');
    ASSERT_FALSE(fb.CMD.ARMPULSE_CMD, 'BtnEmergencyCutOff doit aussi couper le pulse de reamement en cours');
    ASSERT_EQ(fb.STATUS.STATE.STEP, 0, 'BtnEmergencyCutOff ramene immediatement a Step 0');
    ASSERT_EQ(fb.STATUS.DIAG.LASTABORTCAUSE, 16#0001, 'LastAbortCause = CST_ABORT_CUT_IHM (1)');
END_TEST
